Fanuc KAREL source: kc00040.KL

-- PROVISIONAL review KL for V1013-1; original PC SHA256 f452243ec917a2b963816d7bdef30a776930770d8a88fc8b04def8efd8a50c0a
-- Incomplete behavior may be omitted. Consult companion uncertainty JSON. Do not deploy.
PROGRAM KC00040
%NOLOCKGROUP
BEGIN
  -- UNRESOLVED_PC offsets 5-33; opcodes 27,22,22,22,22,31
  -- UNRESOLVED_PC offsets 38-42; opcodes 7F
END KC00040
